(* IEC 61131-3 sources: test-1/plc/exports, 8 files *)

(* ---- E_CellFault.st ---- *)
{attribute 'qualified_only'}
{attribute 'strict'}
TYPE E_CellFault :
(
    NONE := 0,
    INTERLOCK_OPEN := 1,
    LIMIT_CONFLICT := 2,
    EXIT_CONFLICT := 3,
    START_NOT_CLEAR := 4,
    PUSHER_NOT_HOME := 5,
    UNEXPECTED_EXIT := 6,
    FEED_TIMEOUT := 7,
    ACCEPT_TIMEOUT := 8,
    METAL_ROUTE_NOT_IMPLEMENTED := 9,
    INVALID_STATE := 10,
    COUNT_OVERFLOW := 11
) := NONE;
END_TYPE

(* ---- E_CellState.st ---- *)
{attribute 'qualified_only'}
{attribute 'strict'}
TYPE E_CellState :
(
    STOPPED := 0,
    READY := 1,
    FEED := 2,
    ACCEPT := 3,
    EXTEND := 4,  (* Reserved for Stage 3; invalid in this controller. *)
    RETRACT := 5, (* Reserved for Stage 3; invalid in this controller. *)
    FAULT := 6
) := STOPPED;
END_TYPE

(* ---- ST_CellInputs.st ---- *)
TYPE ST_CellInputs :
STRUCT
    start : BOOL := FALSE;
    reset : BOOL := FALSE;
    stop : BOOL := FALSE;
    permissive_ok : BOOL := TRUE; (* Simulation default, not a safety input. *)
    station : BOOL := FALSE;
    metal : BOOL := FALSE;
    accepted : BOOL := FALSE;
    rejected : BOOL := FALSE;
    pusher_home : BOOL := TRUE;
    pusher_extended : BOOL := FALSE;
END_STRUCT
END_TYPE

(* ---- ST_CellOutputs.st ---- *)
TYPE ST_CellOutputs :
STRUCT
    conveyor : BOOL := FALSE;
    extend : BOOL := FALSE;
    alarm : BOOL := FALSE;
    ready : BOOL := FALSE;
END_STRUCT
END_TYPE

(* ---- ST_Stage2Sample.st ---- *)
TYPE ST_Stage2Sample :
STRUCT
    scan : UINT;
    entry_state : E_CellState;
    inputs : ST_CellInputs;
    state : E_CellState;
    fault : E_CellFault;
    outputs : ST_CellOutputs;
    accepted_count : UDINT;
    accepted_seen : BOOL;
    feed_et : TIME;
    accept_et : TIME;
    feed_q : BOOL;
    accept_q : BOOL;
END_STRUCT
END_TYPE

(* ---- FB_ConveyorSorter.st ---- *)
FUNCTION_BLOCK FB_ConveyorSorter
VAR_INPUT
    i : ST_CellInputs;
END_VAR
VAR_OUTPUT
    o : ST_CellOutputs;
    state : E_CellState := E_CellState.STOPPED;
    fault : E_CellFault := E_CellFault.NONE;
    accepted_count : UDINT := 0;
    rejected_count : UDINT := 0; (* Reserved; never incremented in Stage 2. *)
    accepted_seen : BOOL := FALSE;
    start_edge : BOOL;
    reset_edge : BOOL;
    feed_et : TIME;
    accept_et : TIME;
    feed_q : BOOL;
    accept_q : BOOL;
END_VAR
VAR
    startTrigger : R_TRIG;
    resetTrigger : R_TRIG;
    feedTimer : TON;
    acceptTimer : TON;
    scanState : E_CellState;
    clearPath : BOOL;
END_VAR
VAR CONSTANT
    FEED_TIMEOUT : TIME := T#5s;
    ACCEPT_TIMEOUT : TIME := T#3s;
END_VAR

(* IMPLEMENTATION: paste below this line into the ST implementation pane. *)
(* Simulation-only, one call per 20 ms task. No RETAIN or physical addresses. *)
scanState := state;
startTrigger(CLK := i.start);
resetTrigger(CLK := i.reset);
start_edge := startTrigger.Q;
reset_edge := resetTrigger.Q;
clearPath := NOT (i.station OR i.accepted OR i.rejected)
             AND i.pusher_home AND NOT i.pusher_extended;

(* Preserve the first fault. Global checks precede Stop and normal sequence. *)
IF state <> E_CellState.FAULT THEN
    IF NOT i.permissive_ok THEN
        fault := E_CellFault.INTERLOCK_OPEN;
    ELSIF i.pusher_home AND i.pusher_extended THEN
        fault := E_CellFault.LIMIT_CONFLICT;
    ELSIF i.accepted AND i.rejected THEN
        fault := E_CellFault.EXIT_CONFLICT;
    ELSIF (state <> E_CellState.STOPPED) AND (state <> E_CellState.READY)
        AND (state <> E_CellState.FEED) AND (state <> E_CellState.ACCEPT) THEN
        fault := E_CellFault.INVALID_STATE;
    END_IF;
    IF fault <> E_CellFault.NONE THEN
        state := E_CellState.FAULT;
    END_IF;
END_IF;

IF state = E_CellState.FAULT THEN
    (* A new fault must remain observable for its detection scan.
       A Reset edge consumed on that scan cannot also recover it. *)
    IF (scanState = E_CellState.FAULT) AND reset_edge AND NOT i.start AND NOT i.stop
        AND i.permissive_ok AND clearPath THEN
        fault := E_CellFault.NONE;
        state := E_CellState.READY;
    END_IF;
ELSIF i.stop THEN
    state := E_CellState.STOPPED;
ELSE
    CASE state OF
        E_CellState.STOPPED:
            IF reset_edge AND NOT i.start AND clearPath THEN
                state := E_CellState.READY;
            END_IF;
        E_CellState.READY:
            IF start_edge AND NOT i.reset THEN
                IF clearPath THEN
                    state := E_CellState.FEED;
                ELSE
                    fault := E_CellFault.START_NOT_CLEAR;
                    state := E_CellState.FAULT;
                END_IF;
            END_IF;
    END_CASE;
END_IF;

(* Start FEED's TON on the READY -> FEED scan, not one scan later.
   Each TON is called once every scan, including STOPPED/FAULT scans. *)
feedTimer(IN := state = E_CellState.FEED, PT := FEED_TIMEOUT);
IF (scanState = E_CellState.FEED) AND (state = E_CellState.FEED) THEN
    IF feedTimer.Q THEN
        fault := E_CellFault.FEED_TIMEOUT;
        state := E_CellState.FAULT;
    ELSIF NOT i.pusher_home THEN
        fault := E_CellFault.PUSHER_NOT_HOME;
        state := E_CellState.FAULT;
    ELSIF i.accepted OR i.rejected THEN
        fault := E_CellFault.UNEXPECTED_EXIT;
        state := E_CellState.FAULT;
    ELSIF i.station THEN
        IF i.metal THEN
            fault := E_CellFault.METAL_ROUTE_NOT_IMPLEMENTED;
            state := E_CellState.FAULT;
        ELSE
            state := E_CellState.ACCEPT;
        END_IF;
    END_IF;
END_IF;

(* Start ACCEPT's TON on the FEED -> ACCEPT scan. scanState prevents
   evaluating a newly entered phase twice in one scan. *)
acceptTimer(IN := state = E_CellState.ACCEPT, PT := ACCEPT_TIMEOUT);
IF (scanState = E_CellState.ACCEPT) AND (state = E_CellState.ACCEPT) THEN
    IF acceptTimer.Q THEN
        fault := E_CellFault.ACCEPT_TIMEOUT;
        state := E_CellState.FAULT;
    ELSIF NOT i.pusher_home THEN
        fault := E_CellFault.PUSHER_NOT_HOME;
        state := E_CellState.FAULT;
    ELSIF i.rejected THEN
        fault := E_CellFault.UNEXPECTED_EXIT;
        state := E_CellState.FAULT;
    ELSE
        accepted_seen := accepted_seen OR i.accepted;
        IF accepted_seen AND NOT i.accepted AND NOT i.station THEN
            IF accepted_count = UDINT#4294967295 THEN
                fault := E_CellFault.COUNT_OVERFLOW;
                state := E_CellState.FAULT;
            ELSE
                accepted_count := accepted_count + UDINT#1;
                state := E_CellState.READY;
            END_IF;
        END_IF;
    END_IF;
END_IF;

(* Discard incomplete passage memory on completion, Stop or any fault. *)
IF state <> E_CellState.ACCEPT THEN
    accepted_seen := FALSE;
END_IF;
(* Diagnostics show this scan's timer calls; an exited timer resets on
   its next call (next scan). These are not end-state elapsed counters. *)
feed_et := feedTimer.ET;
accept_et := acceptTimer.ET;
feed_q := feedTimer.Q;
accept_q := acceptTimer.Q;

(* Assign every output every scan from the resulting state. *)
o.conveyor := (state = E_CellState.FEED) OR (state = E_CellState.ACCEPT);
o.extend := FALSE;
o.alarm := state = E_CellState.FAULT;
o.ready := (state = E_CellState.READY) AND clearPath;
END_FUNCTION_BLOCK

(* ---- PLC_PRG.st ---- *)
PROGRAM PLC_PRG
VAR
    simInputs : ST_CellInputs; (* Manual watch-list input image. *)
    sorter : FB_ConveyorSorter;
END_VAR

(* IMPLEMENTATION: paste below this line into the ST implementation pane. *)
sorter(i := simInputs);
END_PROGRAM

(* ---- PRG_TestSequence.st ---- *)
PROGRAM PRG_TestSequence
VAR
    (* Set testCase while stopped after an IDE Reset Cold; then Run.
       0 normal + held Start + Stop/Reset/fresh Start; 1 FEED deadline;
       2 ACCEPT deadline; 3 FEED one scan early; 4 ACCEPT one scan early;
       5 reserved EXTEND + Reset; 6 reserved RETRACT + Reset. *)
    testCase : UINT := 0;
    scan : UINT := 0;
    done : BOOL := FALSE;
    sequence_passed : BOOL := FALSE; (* Assertions only, NOT a measured timing PASS. *)
    failed : BOOL := FALSE;
    inputs : ST_CellInputs;
    dut : FB_ConveyorSorter;
    samples : ARRAY[0..300] OF ST_Stage2Sample;
END_VAR

(* IMPLEMENTATION: paste below this line into the ST implementation pane. *)
(* Simulation-only alternative task entry. Never schedule alongside PLC_PRG.
   Boundary cases use nominal scan counts. External timestamped task traces
   are mandatory for timing verdicts; this array has no measured clock. *)
IF NOT done THEN
    inputs.start := scan >= 2;
    inputs.reset := scan = 1;
    inputs.stop := FALSE;
    inputs.permissive_ok := TRUE;
    inputs.station := FALSE;
    inputs.metal := FALSE;
    inputs.accepted := FALSE;
    inputs.rejected := FALSE;
    inputs.pusher_home := TRUE;
    inputs.pusher_extended := FALSE;
    CASE testCase OF
        0:
            inputs.station := (scan >= 3) AND (scan <= 5);
            inputs.accepted := (scan = 4) OR (scan = 5);
            IF scan >= 9 THEN inputs.start := scan >= 12; END_IF;
            inputs.stop := scan = 9;
            inputs.reset := (scan = 1) OR (scan = 10);
        1:
            inputs.station := scan = 252;
        2:
            inputs.station := scan = 3;
            inputs.accepted := (scan >= 4) AND (scan < 153);
        3:
            inputs.station := scan = 251;
            inputs.accepted := scan = 252;
        4:
            inputs.station := scan = 3;
            inputs.accepted := (scan >= 4) AND (scan < 152);
        5, 6:
            inputs.start := FALSE;
            inputs.reset := (scan = 1) OR (scan = 2) OR (scan = 4);
            (* Deliberate test-only state injection before the detection call.
               Never copy this assignment into PLC_PRG or the controller FB. *)
            IF scan = 1 THEN
                IF testCase = 5 THEN
                    dut.state := E_CellState.EXTEND;
                ELSE
                    dut.state := E_CellState.RETRACT;
                END_IF;
            END_IF;
    ELSE
        failed := TRUE;
        done := TRUE;
    END_CASE;

    IF NOT done THEN
        samples[scan].entry_state := dut.state;
        dut(i := inputs);
        samples[scan].scan := scan;
        samples[scan].inputs := inputs;
        samples[scan].state := dut.state;
        samples[scan].fault := dut.fault;
        samples[scan].outputs := dut.o;
        samples[scan].accepted_count := dut.accepted_count;
        samples[scan].accepted_seen := dut.accepted_seen;
        samples[scan].feed_et := dut.feed_et;
        samples[scan].accept_et := dut.accept_et;
        samples[scan].feed_q := dut.feed_q;
        samples[scan].accept_q := dut.accept_q;

        failed := failed OR dut.o.extend OR (dut.accepted_count > 1)
                  OR (dut.rejected_count <> 0);
        IF scan = 0 THEN
            failed := failed OR (dut.state <> E_CellState.STOPPED)
                      OR dut.o.conveyor OR (dut.accepted_count <> 0);
        ELSIF (scan = 1) AND (testCase <= 4) THEN
            failed := failed OR (dut.state <> E_CellState.READY) OR dut.o.conveyor;
        ELSIF (scan = 2) AND (testCase <= 4) THEN
            failed := failed OR (dut.state <> E_CellState.FEED)
                      OR NOT dut.o.conveyor OR (dut.feed_et <> T#0ms);
        END_IF;

        CASE testCase OF
            0:
                IF (scan >= 3) AND (scan <= 5) THEN
                    failed := failed OR (dut.state <> E_CellState.ACCEPT)
                              OR (dut.accepted_count <> 0);
                    IF scan = 3 THEN
                        failed := failed OR (dut.accept_et <> T#0ms) OR dut.accept_q;
                    ELSE
                        failed := failed OR (dut.feed_et <> T#0ms) OR dut.feed_q;
                    END_IF;
                ELSIF (scan >= 6) AND (scan <= 8) THEN
                    failed := failed OR (dut.state <> E_CellState.READY)
                              OR (dut.accepted_count <> 1) OR dut.o.conveyor;
                    IF scan >= 7 THEN
                        failed := failed OR (dut.accept_et <> T#0ms) OR dut.accept_q;
                    END_IF;
                ELSIF scan = 9 THEN
                    failed := failed OR (dut.state <> E_CellState.STOPPED)
                              OR dut.o.conveyor OR (dut.accepted_count <> 1);
                ELSIF (scan = 10) OR (scan = 11) THEN
                    failed := failed OR (dut.state <> E_CellState.READY)
                              OR dut.o.conveyor OR (dut.accepted_count <> 1);
                ELSIF scan >= 12 THEN
                    failed := failed OR (dut.state <> E_CellState.FEED)
                              OR NOT dut.o.conveyor OR (dut.accepted_count <> 1)
                              OR dut.feed_q OR (dut.accept_et <> T#0ms) OR dut.accept_q;
                    IF scan = 12 THEN
                        failed := failed OR (dut.feed_et <> T#0ms);
                    END_IF;
                END_IF;
                done := scan = 13;
            1:
                IF (scan >= 2) AND (scan < 252) THEN
                    failed := failed OR (dut.state <> E_CellState.FEED)
                              OR (dut.accepted_count <> 0);
                ELSIF scan = 252 THEN
                    failed := failed OR (samples[251].state <> E_CellState.FEED)
                              OR samples[251].inputs.station OR NOT inputs.station
                              OR (dut.state <> E_CellState.FAULT)
                              OR (dut.fault <> E_CellFault.FEED_TIMEOUT)
                              OR NOT dut.feed_q OR dut.o.conveyor
                              OR (dut.accepted_count <> 0);
                ELSIF scan = 253 THEN
                    failed := failed OR (dut.state <> E_CellState.FAULT)
                              OR (dut.fault <> E_CellFault.FEED_TIMEOUT)
                              OR dut.feed_q OR (dut.feed_et <> T#0ms)
                              OR dut.o.conveyor OR NOT dut.o.alarm
                              OR (dut.accepted_count <> 0);
                    done := TRUE;
                END_IF;
            2:
                IF (scan >= 3) AND (scan < 153) THEN
                    failed := failed OR (dut.state <> E_CellState.ACCEPT)
                              OR (dut.accepted_count <> 0);
                ELSIF scan = 153 THEN
                    failed := failed OR (samples[152].state <> E_CellState.ACCEPT)
                              OR NOT samples[152].inputs.accepted OR inputs.accepted
                              OR (dut.state <> E_CellState.FAULT)
                              OR (dut.fault <> E_CellFault.ACCEPT_TIMEOUT)
                              OR NOT dut.accept_q OR dut.o.conveyor
                              OR (dut.accepted_count <> 0);
                ELSIF scan = 154 THEN
                    failed := failed OR (dut.state <> E_CellState.FAULT)
                              OR (dut.fault <> E_CellFault.ACCEPT_TIMEOUT)
                              OR dut.accept_q OR (dut.accept_et <> T#0ms)
                              OR dut.o.conveyor OR NOT dut.o.alarm
                              OR (dut.accepted_count <> 0);
                    done := TRUE;
                END_IF;
            3:
                IF (scan >= 2) AND (scan < 251) THEN
                    failed := failed OR (dut.state <> E_CellState.FEED)
                              OR (dut.accepted_count <> 0) OR dut.feed_q;
                ELSIF scan = 251 THEN
                    failed := failed OR (samples[250].state <> E_CellState.FEED)
                              OR (samples[250].accepted_count <> 0)
                              OR samples[250].inputs.station OR NOT inputs.station
                              OR (samples[251].entry_state <> E_CellState.FEED)
                              OR (dut.state <> E_CellState.ACCEPT)
                              OR (dut.accepted_count <> 0) OR dut.feed_q
                              OR (dut.feed_et >= T#5s) OR (dut.accept_et <> T#0ms);
                ELSIF scan = 252 THEN
                    failed := failed OR (dut.state <> E_CellState.ACCEPT)
                              OR NOT inputs.accepted OR NOT dut.accepted_seen
                              OR (dut.accepted_count <> 0)
                              OR dut.feed_q OR (dut.feed_et <> T#0ms);
                ELSIF scan = 253 THEN
                    failed := failed OR (samples[252].accepted_count <> 0)
                              OR NOT samples[252].inputs.accepted OR inputs.accepted
                              OR (dut.state <> E_CellState.READY)
                              OR (dut.accepted_count <> 1) OR dut.o.conveyor;
                    done := TRUE;
                END_IF;
            4:
                IF (scan >= 3) AND (scan < 152) THEN
                    failed := failed OR (dut.state <> E_CellState.ACCEPT)
                              OR (dut.accepted_count <> 0) OR dut.accept_q;
                ELSIF scan = 152 THEN
                    failed := failed OR (samples[151].state <> E_CellState.ACCEPT)
                              OR (samples[151].accepted_count <> 0)
                              OR NOT samples[151].accepted_seen
                              OR NOT samples[151].inputs.accepted
                              OR inputs.accepted OR inputs.station
                              OR (samples[152].entry_state <> E_CellState.ACCEPT)
                              OR (dut.state <> E_CellState.READY)
                              OR dut.accept_q OR (dut.accept_et >= T#3s)
                              OR (dut.accepted_count <> 1) OR dut.o.conveyor;
                ELSIF scan = 153 THEN
                    failed := failed OR (dut.state <> E_CellState.READY)
                              OR (dut.accepted_count <> 1) OR dut.o.conveyor
                              OR dut.accept_q OR (dut.accept_et <> T#0ms);
                    done := TRUE;
                END_IF;
            5, 6:
                IF (scan >= 1) AND (scan <= 3) THEN
                    failed := failed OR (dut.state <> E_CellState.FAULT)
                              OR (dut.fault <> E_CellFault.INVALID_STATE)
                              OR NOT dut.o.alarm OR dut.o.ready;
                ELSIF scan >= 4 THEN
                    failed := failed OR (dut.state <> E_CellState.READY)
                              OR (dut.fault <> E_CellFault.NONE)
                              OR dut.o.alarm OR NOT dut.o.ready;
                END_IF;
                failed := failed OR dut.o.conveyor OR (dut.accepted_count <> 0)
                          OR dut.feed_q OR dut.accept_q;
                done := scan = 5;
        END_CASE;
        IF scan = 300 THEN
            failed := TRUE;
            done := TRUE;
        END_IF;
        sequence_passed := done AND NOT failed;
        IF NOT done THEN scan := scan + 1; END_IF;
    END_IF;
END_IF;
(* The runner stops calling its private DUT when done. Timeout modes include
   the following reset-diagnostic scan, but NOT fault recovery. S2-20 requires
   a separate continuous recovery trace. No runtime evidence exists until run. *)
END_PROGRAM
